(* PLC project a.project, CODESYS CODESYS V3.5 SP17 Patch 3 *)
(* stored: creationDateTime 2026-10-19T00:00:00, modificationDateTime 2026-10-19T00:00:00 *)

FUNCTION_BLOCK FB_Act
VAR
    n : INT;
END_VAR

            ActInc();

          

ACTION ActInc:
                n := n + 1;

              
END_ACTION
END_FUNCTION_BLOCK
